FUNCTION_BLOCK "FB_StlC_054"   // FB70, STL
TITLE = STL call UPPER_BOUND
{ S7_Optimized_Access := 'TRUE' }
VERSION : 0.1
   VAR_INPUT
      "a" : Bool;
      i1 : Int;
      i2 : Int;
      di1 : DInt;
      r1 : Real;
      w1 : Word;
      dw1 : DWord;
      b1 : Byte;
      u1 : UInt;
      ud1 : UDInt;
   END_VAR
   VAR_OUTPUT
      q : Bool;
      io : Int;
      dio : DInt;
      ro : Real;
      wo : Word;
      dwo : DWord;
      bo : Byte;
      udo : UDInt;
   END_VAR
   VAR_IN_OUT
      v : Variant;
      arrs : Array[*] of Int;
      pos : DInt;
   END_VAR
   VAR
      src : Array[0..9] of Int;
      dst : Array[0..9] of Int;
      bits : Array[0..31] of Bool;
      bytes : Array[0..9] of Byte;
      err : ErrorStruct;
      rt : LReal;
      tim : IEC_TIMER;
      words : Array[0..3] of Word;
   END_VAR
BEGIN

REGION Network 1: 054 UPPER_BOUND
         CALL  UPPER_BOUND
         ( ARR := #arrs,
           DIM := #ud1,
           OUT := #dio
         );
END_REGION
END_FUNCTION_BLOCK

FUNCTION_BLOCK "FB_StlC_057"   // FB71, STL
TITLE = STL call FILL
{ S7_Optimized_Access := 'TRUE' }
VERSION : 0.1
   VAR_INPUT
      "a" : Bool;
      i1 : Int;
      i2 : Int;
      di1 : DInt;
      r1 : Real;
      w1 : Word;
      dw1 : DWord;
      b1 : Byte;
      u1 : UInt;
      ud1 : UDInt;
   END_VAR
   VAR_OUTPUT
      q : Bool;
      io : Int;
      dio : DInt;
      ro : Real;
      wo : Word;
      dwo : DWord;
      bo : Byte;
      udo : UDInt;
   END_VAR
   VAR_IN_OUT
      v : Variant;
      arrs : Array[*] of Int;
      pos : DInt;
   END_VAR
   VAR
      src : Array[0..9] of Int;
      dst : Array[0..9] of Int;
      bits : Array[0..31] of Bool;
      bytes : Array[0..9] of Byte;
      err : ErrorStruct;
      rt : LReal;
      tim : IEC_TIMER;
      words : Array[0..3] of Word;
   END_VAR
BEGIN

REGION Network 1: 057 FILL
         CALL  FILL
         ( BVAL    := #v,
           RET_VAL := #io,
           BLK     := #v
         );
END_REGION
END_FUNCTION_BLOCK

FUNCTION_BLOCK "FB_StlC_013"   // FB72, STL
TITLE = STL call EQ_Type
{ S7_Optimized_Access := 'TRUE' }
VERSION : 0.1
   VAR_INPUT
      "a" : Bool;
      i1 : Int;
      i2 : Int;
      di1 : DInt;
      r1 : Real;
      w1 : Word;
      dw1 : DWord;
      b1 : Byte;
      u1 : UInt;
      ud1 : UDInt;
   END_VAR
   VAR_OUTPUT
      q : Bool;
      io : Int;
      dio : DInt;
      ro : Real;
      wo : Word;
      dwo : DWord;
      bo : Byte;
      udo : UDInt;
   END_VAR
   VAR_IN_OUT
      v : Variant;
      arrs : Array[*] of Int;
      pos : DInt;
   END_VAR
   VAR
      src : Array[0..9] of Int;
      dst : Array[0..9] of Int;
      bits : Array[0..31] of Bool;
      bytes : Array[0..9] of Byte;
      err : ErrorStruct;
      rt : LReal;
      tim : IEC_TIMER;
      words : Array[0..3] of Word;
   END_VAR
BEGIN

REGION Network 1: 013 EQ_Type
         CALL  EQ_Type
         ( IN1     := #v,
           IN2     := #i1,
           Ret_Val := #q
         );
END_REGION
END_FUNCTION_BLOCK

FUNCTION_BLOCK "FB_StlC_014"   // FB73, STL
TITLE = STL call NE_Type
{ S7_Optimized_Access := 'TRUE' }
VERSION : 0.1
   VAR_INPUT
      "a" : Bool;
      i1 : Int;
      i2 : Int;
      di1 : DInt;
      r1 : Real;
      w1 : Word;
      dw1 : DWord;
      b1 : Byte;
      u1 : UInt;
      ud1 : UDInt;
   END_VAR
   VAR_OUTPUT
      q : Bool;
      io : Int;
      dio : DInt;
      ro : Real;
      wo : Word;
      dwo : DWord;
      bo : Byte;
      udo : UDInt;
   END_VAR
   VAR_IN_OUT
      v : Variant;
      arrs : Array[*] of Int;
      pos : DInt;
   END_VAR
   VAR
      src : Array[0..9] of Int;
      dst : Array[0..9] of Int;
      bits : Array[0..31] of Bool;
      bytes : Array[0..9] of Byte;
      err : ErrorStruct;
      rt : LReal;
      tim : IEC_TIMER;
      words : Array[0..3] of Word;
   END_VAR
BEGIN

REGION Network 1: 014 NE_Type
         CALL  NE_Type
         ( IN1     := #v,
           IN2     := #i1,
           Ret_Val := #q
         );
END_REGION
END_FUNCTION_BLOCK

FUNCTION_BLOCK "FB_StlC_015"   // FB74, STL
TITLE = STL call EQ_ElemType
{ S7_Optimized_Access := 'TRUE' }
VERSION : 0.1
   VAR_INPUT
      "a" : Bool;
      i1 : Int;
      i2 : Int;
      di1 : DInt;
      r1 : Real;
      w1 : Word;
      dw1 : DWord;
      b1 : Byte;
      u1 : UInt;
      ud1 : UDInt;
   END_VAR
   VAR_OUTPUT
      q : Bool;
      io : Int;
      dio : DInt;
      ro : Real;
      wo : Word;
      dwo : DWord;
      bo : Byte;
      udo : UDInt;
   END_VAR
   VAR_IN_OUT
      v : Variant;
      arrs : Array[*] of Int;
      pos : DInt;
   END_VAR
   VAR
      src : Array[0..9] of Int;
      dst : Array[0..9] of Int;
      bits : Array[0..31] of Bool;
      bytes : Array[0..9] of Byte;
      err : ErrorStruct;
      rt : LReal;
      tim : IEC_TIMER;
      words : Array[0..3] of Word;
   END_VAR
BEGIN

REGION Network 1: 015 EQ_ElemType
         CALL  EQ_ElemType
         ( IN1     := #v,
           IN2     := #i1,
           Ret_Val := #q
         );
END_REGION
END_FUNCTION_BLOCK

FUNCTION_BLOCK "FB_StlC_016"   // FB75, STL
TITLE = STL call NE_ElemType
{ S7_Optimized_Access := 'TRUE' }
VERSION : 0.1
   VAR_INPUT
      "a" : Bool;
      i1 : Int;
      i2 : Int;
      di1 : DInt;
      r1 : Real;
      w1 : Word;
      dw1 : DWord;
      b1 : Byte;
      u1 : UInt;
      ud1 : UDInt;
   END_VAR
   VAR_OUTPUT
      q : Bool;
      io : Int;
      dio : DInt;
      ro : Real;
      wo : Word;
      dwo : DWord;
      bo : Byte;
      udo : UDInt;
   END_VAR
   VAR_IN_OUT
      v : Variant;
      arrs : Array[*] of Int;
      pos : DInt;
   END_VAR
   VAR
      src : Array[0..9] of Int;
      dst : Array[0..9] of Int;
      bits : Array[0..31] of Bool;
      bytes : Array[0..9] of Byte;
      err : ErrorStruct;
      rt : LReal;
      tim : IEC_TIMER;
      words : Array[0..3] of Word;
   END_VAR
BEGIN

REGION Network 1: 016 NE_ElemType
         CALL  NE_ElemType
         ( IN1     := #v,
           IN2     := #i1,
           Ret_Val := #q
         );
END_REGION
END_FUNCTION_BLOCK

FUNCTION_BLOCK "FB_StlC_018"   // FB76, STL
TITLE = STL call NOT_NULL
{ S7_Optimized_Access := 'TRUE' }
VERSION : 0.1
   VAR_INPUT
      "a" : Bool;
      i1 : Int;
      i2 : Int;
      di1 : DInt;
      r1 : Real;
      w1 : Word;
      dw1 : DWord;
      b1 : Byte;
      u1 : UInt;
      ud1 : UDInt;
   END_VAR
   VAR_OUTPUT
      q : Bool;
      io : Int;
      dio : DInt;
      ro : Real;
      wo : Word;
      dwo : DWord;
      bo : Byte;
      udo : UDInt;
   END_VAR
   VAR_IN_OUT
      v : Variant;
      arrs : Array[*] of Int;
      pos : DInt;
   END_VAR
   VAR
      src : Array[0..9] of Int;
      dst : Array[0..9] of Int;
      bits : Array[0..31] of Bool;
      bytes : Array[0..9] of Byte;
      err : ErrorStruct;
      rt : LReal;
      tim : IEC_TIMER;
      words : Array[0..3] of Word;
   END_VAR
BEGIN

REGION Network 1: 018 NOT_NULL
         CALL  NOT_NULL
         ( OPERAND := #v,
           Ret_Val := #q
         );
END_REGION
END_FUNCTION_BLOCK

FUNCTION_BLOCK "FB_StlC_019"   // FB77, STL
TITLE = STL call IS_ARRAY
{ S7_Optimized_Access := 'TRUE' }
VERSION : 0.1
   VAR_INPUT
      "a" : Bool;
      i1 : Int;
      i2 : Int;
      di1 : DInt;
      r1 : Real;
      w1 : Word;
      dw1 : DWord;
      b1 : Byte;
      u1 : UInt;
      ud1 : UDInt;
   END_VAR
   VAR_OUTPUT
      q : Bool;
      io : Int;
      dio : DInt;
      ro : Real;
      wo : Word;
      dwo : DWord;
      bo : Byte;
      udo : UDInt;
   END_VAR
   VAR_IN_OUT
      v : Variant;
      arrs : Array[*] of Int;
      pos : DInt;
   END_VAR
   VAR
      src : Array[0..9] of Int;
      dst : Array[0..9] of Int;
      bits : Array[0..31] of Bool;
      bytes : Array[0..9] of Byte;
      err : ErrorStruct;
      rt : LReal;
      tim : IEC_TIMER;
      words : Array[0..3] of Word;
   END_VAR
BEGIN

REGION Network 1: 019 IS_ARRAY
         CALL  IS_ARRAY
         ( OPERAND := #v,
           Ret_Val := #q
         );
END_REGION
END_FUNCTION_BLOCK

FUNCTION_BLOCK "FB_StlC_036"   // FB78, STL
TITLE = STL call GATHER_BLK
{ S7_Optimized_Access := 'TRUE' }
VERSION : 0.1
   VAR_INPUT
      "a" : Bool;
      i1 : Int;
      i2 : Int;
      di1 : DInt;
      r1 : Real;
      w1 : Word;
      dw1 : DWord;
      b1 : Byte;
      u1 : UInt;
      ud1 : UDInt;
   END_VAR
   VAR_OUTPUT
      q : Bool;
      io : Int;
      dio : DInt;
      ro : Real;
      wo : Word;
      dwo : DWord;
      bo : Byte;
      udo : UDInt;
   END_VAR
   VAR_IN_OUT
      v : Variant;
      arrs : Array[*] of Int;
      pos : DInt;
   END_VAR
   VAR
      src : Array[0..9] of Int;
      dst : Array[0..9] of Int;
      bits : Array[0..31] of Bool;
      bytes : Array[0..9] of Byte;
      err : ErrorStruct;
      rt : LReal;
      tim : IEC_TIMER;
      words : Array[0..3] of Word;
   END_VAR
BEGIN

REGION Network 1: 036 GATHER_BLK
         CALL  GATHER_BLK
         ( IN        := #bits[0],
           COUNT_OUT := #u1,
           OUT       := #words[0]
         );
END_REGION
END_FUNCTION_BLOCK

FUNCTION_BLOCK "FB_StlC_055"   // FB79, STL
TITLE = STL call BLKMOV
{ S7_Optimized_Access := 'FALSE' }
VERSION : 0.1
   VAR_OUTPUT
      io : Int;
   END_VAR
BEGIN

REGION Network 1: 055 BLKMOV
         CALL  BLKMOV
         ( SRCBLK  := "DB_Arr"."a",
           RET_VAL := #io,
           DSTBLK  := "DB_Arr"."b"
         );
END_REGION

REGION Network 2: 056 UBLKMOV
         CALL  UBLKMOV
         ( SRCBLK  := "DB_Arr"."a",
           RET_VAL := #io,
           DSTBLK  := "DB_Arr"."b"
         );
END_REGION
END_FUNCTION_BLOCK

FUNCTION_BLOCK "FB_StlC_060"   // FB85, STL
TITLE = STL call VARIANT_TO_DB_ANY
{ S7_Optimized_Access := 'TRUE' }
VERSION : 0.1
   VAR_OUTPUT
      io : Int;
   END_VAR
   VAR_IN_OUT
      v : Variant;
   END_VAR
   VAR_TEMP
      dba : DB_ANY;
   END_VAR
BEGIN

REGION Network 1: 060 VARIANT_TO_DB_ANY
         CALL  VARIANT_TO_DB_ANY
         ( in      := #v,
           Ret_Val := #dba,
           err     := #io
         );
END_REGION

REGION Network 2: 061 DB_ANY_TO_VARIANT
         CALL  DB_ANY_TO_VARIANT
         ( in      := #dba,
           Ret_Val := #v,
           err     := #io
         );
END_REGION
END_FUNCTION_BLOCK

FUNCTION_BLOCK "FB_StlC_037"   // FB86, STL
TITLE = STL call ReadFromArrayDB
{ S7_Optimized_Access := 'TRUE' }
VERSION : 0.1
   VAR_INPUT
      di1 : DInt;
   END_VAR
   VAR_OUTPUT
      io : Int;
   END_VAR
   VAR
      val : Int;
   END_VAR
BEGIN

REGION Network 1: 037 ReadFromArrayDB
         CALL  ReadFromArrayDB
         ( db      := "ArrDB",
           index   := #di1,
           Ret_Val := #io,
           value   := #val
         );
END_REGION

REGION Network 2: 038 WriteToArrayDB
         CALL  WriteToArrayDB
         ( db      := "ArrDB",
           index   := #di1,
           value   := #val,
           Ret_Val := #io
         );
END_REGION
END_FUNCTION_BLOCK

FUNCTION_BLOCK "FB_StlC_029"   // FB87, STL
TITLE = STL call MOVE_BLK_VARIANT
{ S7_Optimized_Access := 'TRUE' }
VERSION : 0.1
   VAR_INPUT
      cnt : UDInt;
      si : DInt;
      di : DInt;
   END_VAR
   VAR_OUTPUT
      io : Int;
   END_VAR
   VAR_IN_OUT
      src : Variant;
      dst : Variant;
   END_VAR
BEGIN

REGION Network 1: 029 MOVE_BLK_VARIANT
         CALL  MOVE_BLK_VARIANT
         ( SRC        := #src,
           COUNT      := #cnt,
           SRC_INDEX  := #si,
           DEST_INDEX := #di,
           Ret_Val    := #io,
           DEST       := #dst
         );
END_REGION
END_FUNCTION_BLOCK

FUNCTION_BLOCK "FB_StlC_008"   // FB88, STL
TITLE = STL call PRESET_TIMER
{ S7_Optimized_Access := 'TRUE' }
VERSION : 0.1
   VAR
      t1 : IEC_TIMER;
   END_VAR
BEGIN

REGION Network 1: 008 PRESET_TIMER
         CALL  PRESET_TIMER
         ( PT      := T#2S,
           "TIMER" := #t1
         );
END_REGION
END_FUNCTION_BLOCK

FUNCTION_BLOCK "FB_StlC_012"   // FB89, STL
TITLE = STL call CompType
{ S7_Optimized_Access := 'TRUE' }
VERSION : 0.1
   VAR_OUTPUT
      "b" : Bool;
   END_VAR
   VAR
      a1 : Array[0..3] of Int;
      a2 : Array[0..3] of Int;
   END_VAR
BEGIN

REGION Network 1: 012 CompType
         CALL  CompType
         ( IN1 := #a1,
           IN2 := #a2,
           OUT := #"b"
         );
END_REGION
END_FUNCTION_BLOCK

FUNCTION_BLOCK "FB_StlC_020"   // FB90, STL
TITLE = STL call EQ_TypeOfDB
{ S7_Optimized_Access := 'TRUE' }
VERSION : 0.1
   VAR_INPUT
      dba : DB_ANY;
   END_VAR
   VAR_OUTPUT
      "b" : Bool;
   END_VAR
BEGIN

REGION Network 1: 020 EQ_TypeOfDB
         CALL  EQ_TypeOfDB
         ( IN1     := #dba,
           IN2     := "IEC_TIMER",
           Ret_Val := #"b"
         );
END_REGION
END_FUNCTION_BLOCK

FUNCTION_BLOCK "FB_StlC_021"   // FB91, STL
TITLE = STL call NE_TypeOfDB
{ S7_Optimized_Access := 'TRUE' }
VERSION : 0.1
   VAR_INPUT
      dba : DB_ANY;
   END_VAR
   VAR_OUTPUT
      "b" : Bool;
   END_VAR
BEGIN

REGION Network 1: 021 NE_TypeOfDB
         CALL  NE_TypeOfDB
         ( IN1     := #dba,
           IN2     := "IEC_TIMER",
           Ret_Val := #"b"
         );
END_REGION
END_FUNCTION_BLOCK

FUNCTION_BLOCK "FB_StlC_039"   // FB92, STL
TITLE = STL call ReadFromArrayDBL
{ S7_Optimized_Access := 'TRUE' }
VERSION : 0.1
   VAR_INPUT
      req : Bool;
      di1 : DInt;
      dba : DB_ANY;
   END_VAR
   VAR_OUTPUT
      busy : Bool;
      done : Bool;
      err : Int;
   END_VAR
   VAR
      val : Int;
      inst : ReadFromArrayDBL;
   END_VAR
BEGIN

REGION Network 1: 039 ReadFromArrayDBL
         CALL  #inst
         ( req   := #req,
           db    := #dba,
           index := #di1,
           busy  := #busy,
           done  := #done,
           error := #err,
           value := #val
         );
END_REGION
END_FUNCTION_BLOCK

FUNCTION_BLOCK "FB_StlC_040"   // FB93, STL
TITLE = STL call WriteToArrayDBL
{ S7_Optimized_Access := 'TRUE' }
VERSION : 0.1
   VAR_INPUT
      req : Bool;
      di1 : DInt;
      dba : DB_ANY;
   END_VAR
   VAR_OUTPUT
      busy : Bool;
      done : Bool;
      err : Int;
   END_VAR
   VAR
      val : Int;
      inst : WriteToArrayDBL;
   END_VAR
BEGIN

REGION Network 1: 040 WriteToArrayDBL
         CALL  #inst
         ( req   := #req,
           db    := #dba,
           index := #di1,
           value := #val,
           busy  := #busy,
           done  := #done,
           error := #err
         );
END_REGION
END_FUNCTION_BLOCK

FUNCTION_BLOCK "FB_StlC_075"   // FB94, STL
TITLE = STL call DRUM
{ S7_Optimized_Access := 'TRUE' }
VERSION : 0.1
   VAR_INPUT
      req : Bool;
      ev : Bool;
   END_VAR
   VAR_OUTPUT
      "b" : Bool;
      q : Bool;
      ow : Word;
      ec : Word;
   END_VAR
   VAR
      drm : DRUM;
   END_VAR
BEGIN

REGION Network 1: 075 DRUM
         CALL  #drm
         ( RESET    := #req,
           JOG      := #ev,
           DRUM_EN  := #req,
           LST_STEP := B#16#10,
           EVENT1   := #ev,
           EVENT2   := #ev,
           EVENT3   := ,
           EVENT4   := ,
           EVENT5   := ,
           EVENT6   := ,
           EVENT7   := ,
           EVENT8   := ,
           EVENT9   := ,
           EVENT10  := ,
           EVENT11  := ,
           EVENT12  := ,
           EVENT13  := ,
           EVENT14  := ,
           EVENT15  := ,
           EVENT16  := ,
           OUT1     := #"b",
           OUT2     := ,
           OUT3     := ,
           OUT4     := ,
           OUT5     := ,
           OUT6     := ,
           OUT7     := ,
           OUT8     := ,
           OUT9     := ,
           OUT10    := ,
           OUT11    := ,
           OUT12    := ,
           OUT13    := ,
           OUT14    := ,
           OUT15    := ,
           OUT16    := ,
           Q        := #q,
           OUT_WORD := #ow,
           ERR_CODE := #ec
         );
END_REGION
END_FUNCTION_BLOCK

FUNCTION "FC_Stl" : Void   // FC1, STL
TITLE = STL test FC
{ S7_Optimized_Access := 'TRUE' }
VERSION : 0.1
   VAR_INPUT
      "a" : Bool;
      "b" : Bool;
      x : Int;
      y : Int;
   END_VAR
   VAR_OUTPUT
      q : Bool;
      sum : Int;
   END_VAR
   VAR_TEMP
      t : Int;
   END_VAR
BEGIN

REGION Network 1: Bit logic
   // Network comment line 1
         A     #"a";  // and a
         AN    #"b";
         =     #q;
END_REGION

REGION Network 2: Arithmetic
         L     #x;
         L     #y;
         +I;
         T     #t;

         L     #t;
         L     0;
         >I;
         JC    M001;
         L     0;
         T     #t;
   M001: L     #t;
         T     #sum;
END_REGION
END_FUNCTION

FUNCTION "FC_StlNoPar" : Void   // FC2, STL
{ S7_Optimized_Access := 'FALSE' }
VERSION : 0.1
BEGIN

REGION Network 1
         NOP   0;
END_REGION
END_FUNCTION

FUNCTION "FC_StlPar" : Void   // FC3, STL
{ S7_Optimized_Access := 'TRUE' }
VERSION : 0.1
   VAR_INPUT
      x : Int;
      y : Int;
   END_VAR
   VAR_OUTPUT
      q : Bool;
      r : Int;
   END_VAR
BEGIN

REGION Network 1
         L     #x;
         L     #y;
         +I;
         T     #r;
         >I;
         =     #q;
END_REGION
END_FUNCTION

ORGANIZATION_BLOCK "Main"   // OB1, LAD, ProgramCycle
TITLE = "Main Program Sweep (Cycle)"
{ S7_Optimized_Access := 'TRUE' }
VERSION : 0.1
   VAR_INPUT
      Initial_Call : Bool;   // Initial call of this OB
      Remanence : Bool;   // =True, if remanent data are available
   END_VAR
BEGIN
END_ORGANIZATION_BLOCK